(* IEC 61131-3 sources: TcView/src/tests/regression/golden/converter, 2 files *)

(* ---- E_DeviceMode.st ---- *)
TYPE E_DeviceMode :
{attribute 'qualified_only'}
(
    Auto := 0,
    Manual := 1,
    SemiAuto := 2
);
END_TYPE

(* ---- ST_CiA402_Drive_PDO.st ---- *)
TYPE ST_CiA402_Drive_PDO :
STRUCT
    ControlWord    : WORD;
    VelocityTarget : INT;
    StatusWord     : WORD;
    VelocityActual : INT;
    FaultCode      : WORD;
END_STRUCT
END_TYPE
